// TIA Portal V20 export
DATA_BLOCK "T2_Datos"   // DB40921
{ S7_Optimized_Access := 'TRUE' }
AUTHOR : IA
FAMILY : PRUEBA
VERSION : 0.1
// Prueba IA 2: datos de las pruebas
// stored: AutoNumber false
   VAR
      Falso : Bool := false;   // Siempre FALSE
      Verdadero : Bool := true;   // Siempre TRUE
      Mem_Set : Bool;
      Mem_Reset : Bool;
      Mem_Flanco : Bool;
      Int_5 : Int := 5;   // Constante 5
      Word_1234 : Word := 16#1234;   // Constante 16#1234
      Real_2_5 : Real := 2.5;   // Constante 2.5
      DInt_100 : DInt := 100;   // Constante 100
      Move_1 : Int;
      Move_2a : Int;
      Move_2b : Int;
      Swap_Out : Word;
      Conv_Real : Real;
      Str_Hola : String;
      Len_Hola : Int;
      Udt_A : "T2_UDT_Padre";   // Origen de Serialize
      Udt_B : "T2_UDT_Padre";   // Destino de Deserialize
      Buffer : Array[0..99] of Byte;
      PosS : DInt;
      PosD : DInt;
      Ret_Ser : Int;
      Ret_Des : Int;
      Calc_Out : Int;
      Add_Out : Int;
      Sub_Out : Int;
      Concat_Out : String;
      Len_Concat : Int;
      P_Val : UInt := 1;   // Posición VAL_STRG
      P_Strg : UInt := 1;   // Posición STRG_VAL
      Val_Str : String;
      Strg_Int : Int;
      Str_20 : String[20];
      MaxLen_Out : Int;
      Str_Xyz : String := 'XYZ';   // Constante 'XYZ'
      Cnt_Chars : UInt;
      Chars : Array[0..9] of Char;
      Tmr : IEC_TIMER;   // TON de T2_Tiempo
      Rd_Ret : Int;
      Rd_Dtl : DTL;
      Doble_Out : Int;
      FbKop_Q : Bool;
      SclFb_Suma : Int;
      Lista : Array[0..2] of "T2_UDT_Hijo";   // Array de UDT (SCL)
   END_VAR
BEGIN
END_DATA_BLOCK
